Fanuc KAREL source: kd00046.KL

-- PROVISIONAL review KL for V940-1; original PC SHA256 fe3808f8fe489fdb3473c547f53e24bead5962d4d4e155b48fd27dc9f9c7a0f2
-- Incomplete behavior may be omitted. Consult companion uncertainty JSON. Do not deploy.
PROGRAM KD00046
%NOLOCKGROUP
VAR
  I : INTEGER
  J : INTEGER
  B : BOOLEAN
  R : REAL
  S : STRING[80]
-- UNRESOLVED_DECL V type=000013
BEGIN
  -- V9_ZERO_TABLE_METADATA_HINT layout=0001; no indexed target words; source/name/runtime held
  -- UNRESOLVED_PC offsets 5-20; opcodes 2E,22,32,35
  -- UNRESOLVED_PC offsets 25-41; opcodes 01,49,0A,82,0B
  -- UNRESOLVED_PC offsets 46-50; opcodes 7F
END KD00046
